Fanuc KAREL source: ko00040.KL

-- PROVISIONAL review KL for V1013-1; original PC SHA256 0e973b5086d021e4e88f56952392698b4dfa6b280ef0f977d56a9b456fbd8537
-- Incomplete behavior may be omitted. Consult companion uncertainty JSON. Do not deploy.
PROGRAM KO00040
%NOLOCKGROUP
BEGIN
  -- UNRESOLVED_PC offsets 5-12; opcodes 9D,23
  -- UNRESOLVED_PC offsets 17-69; opcodes 27,27,49,7E,AD,27,49,7E,AD,22,31,7E,4A
  -- UNRESOLVED_PC offsets 74-78; opcodes 7F
END KO00040
